Fanuc KAREL source: kt00098.KL

-- PROVISIONAL review KL for V940-1; original PC SHA256 85b9152d772b8e04fe6bec18f7c8fb4d7ee83d6b6cb406d0b7f61f4a0d9d041d
-- Incomplete behavior may be omitted. Consult companion uncertainty JSON. Do not deploy.
PROGRAM KT00098
%NOLOCKGROUP
VAR
  I1 : INTEGER
  I2 : INTEGER
  OUT : REAL
BEGIN
  -- V9_ZERO_TABLE_METADATA_HINT layout=0001; no indexed target words; source/name/runtime held
  -- UNRESOLVED_PC offsets 5-16; opcodes 2E,23
  -- UNRESOLVED_PC offsets 21-32; opcodes 2E,23
  -- UNRESOLVED_PC offsets 37-48; opcodes 2E,23
  -- UNRESOLVED_PC offsets 53-64; opcodes 2E,23
  -- UNRESOLVED_PC offsets 69-92; opcodes 21,21,64,29,64,29,6C,23
  -- UNRESOLVED_PC offsets 97-101; opcodes 7F
END KT00098
